{attribute 'qualified_only'}
{attribute 'strict'}
TYPE E_CoreProt :
(
	None		:= 0,	// 기본 보호 아님 (모듈 규칙)
	PcsFault	:= 1,
	PcsComm		:= 2,
	BatFault	:= 3,
	BatComm		:= 4,
	PccInvalid	:= 5	// 접속점 계측 무효
) INT;
END_TYPE

(* stored: Version 1.1.0.1, ProductVersion 3.1.4024.15
   DUT E_CoreProt: Id {2b4537cf-f903-44ea-9446-e31c69fe7bad} *)
